FUNCTION_BLOCK FB_LanguageManager
VAR_INPUT
END_VAR
VAR_OUTPUT
END_VAR
VAR
END_VAR

END_FUNCTION_BLOCK

(* stored: Version 1.1.0.1, ProductVersion 3.1.4024.15
   POU FB_LanguageManager: Id {321c985c-8408-4128-9e43-8b0b78bb10a1}, SpecialFunc None *)
